{attribute 'call_after_init'}
FUNCTION_BLOCK FB_ConveyorBase
VAR_INPUT
    enable : BOOL := TRUE;
    start : BOOL;
    reset : BOOL;
    blocked : BOOL;
    BlockTimeout : TIME := T#300ms;
    StartDelay : TIME := T#100ms;
END_VAR
VAR_OUTPUT
    state : E_ConveyorState := E_ConveyorState.Stopped;
    id : DINT;
    running : BOOL;
    actualSpeed : LREAL;
    ready : BOOL;
    initTrace : DINT;
    baseInitCount : DINT;
    afterInitCount : DINT;
END_VAR
VAR
    config : REFERENCE TO ST_ConveyorConfig;
    startTimer : TON;
    blockTimer : TON;
    factor : LREAL;
END_VAR

EvaluateState();
UpdateOutputs();

METHOD PUBLIC FB_init : BOOL
VAR_INPUT
    bInitRetains : BOOL;
    bInCopyCode : BOOL;
    conveyorId : DINT;
    sharedConfig : REFERENCE TO ST_ConveyorConfig;
END_VAR
id := conveyorId;
config REF= sharedConfig;
baseInitCount := baseInitCount + 1;
initTrace := initTrace * 10 + 1;
FB_init := TRUE;
END_METHOD

PROPERTY PUBLIC SpeedFactor : LREAL
GET
SpeedFactor := factor;
END_GET
SET
factor := SpeedFactor;
(* Instrumentation of this example's setup order. *)
initTrace := initTrace * 10 + 3;
END_SET
END_PROPERTY

{attribute 'call_after_init'}
METHOD PUBLIC AfterInit
afterInitCount := afterInitCount + 1;
initTrace := initTrace * 10 + 4;
END_METHOD

ACTION EvaluateState:
IF state = E_ConveyorState.Fault THEN
    IF reset AND NOT blocked THEN
        state := E_ConveyorState.Stopped;
    END_IF;
ELSIF NOT (ready AND enable AND start AND_THEN config.enabled) THEN
    state := E_ConveyorState.Stopped;
ELSIF state = E_ConveyorState.Stopped THEN
    state := E_ConveyorState.Starting;
END_IF;

startTimer(IN := state = E_ConveyorState.Starting OR state = E_ConveyorState.Running,
           PT := StartDelay);
blockTimer(IN := (state = E_ConveyorState.Starting OR state = E_ConveyorState.Running)
                 AND blocked, PT := BlockTimeout);

IF (state = E_ConveyorState.Starting OR state = E_ConveyorState.Running)
   AND blockTimer.Q THEN
    state := E_ConveyorState.Fault;
ELSIF state = E_ConveyorState.Starting AND startTimer.Q THEN
    state := E_ConveyorState.Running;
END_IF;
END_ACTION

ACTION UpdateOutputs:
running := state = E_ConveyorState.Running;
IF running THEN
    actualSpeed := config.speed * factor;
ELSE
    actualSpeed := 0.0;
END_IF;
END_ACTION

END_FUNCTION_BLOCK

(* stored: Version 1.1.0.1, ProductVersion 3.1
   Action EvaluateState: Id {dea59cf8-b235-40a5-ade5-d13ddf675f54}
   Action UpdateOutputs: Id {ce6bf028-987a-4b03-be5a-edcfb7c6faa5} *)
